(* IEC 61131-3 sources: stdmachine/plc/src/07_Tests, 6 files *)

(* ---- FB_AlarmManagerTest.st ---- *)
// Tests du gestionnaire d'alarmes (docs/04 § 10, docs/14 § 5)
FUNCTION_BLOCK FB_AlarmManagerTest EXTENDS TcUnit.FB_TestSuite
VAR
    stBuf : ST_AlarmBuffer;
END_VAR

RaiseTwiceOnce();
ClearedUnackedClosesOnAck();
LatchedEventClosesOnAck();
InfoClosesAtOnce();
AckedConditionClosesOnClear();

METHOD PRIVATE RaiseTwiceOnce
VAR
    fb : FB_AlarmManager;
END_VAR
TEST('RaiseTwiceOnce');
MEMSET(ADR(stBuf), 0, SIZEOF(stBuf));
fb.Bind(stBuf);
fb.Raise(1001, 101, 5, E_Severity.StationFault);
fb.Raise(1001, 101, 6, E_Severity.StationFault);
AssertEquals_UINT(Expected := 1, Actual := stBuf.nActive, Message := 'Une seule alarme pour la meme cle');
AssertEquals_UINT(Expected := 1, Actual := stBuf.aActive[1].nRepeat, Message := 'Repetition comptee');
AssertEquals_UDINT(Expected := 6, Actual := stBuf.aActive[1].nSubCode, Message := 'Sous-code mis a jour');
TEST_FINISHED();
END_METHOD

METHOD PRIVATE ClearedUnackedClosesOnAck
VAR
    fb : FB_AlarmManager;
END_VAR
TEST('ClearedUnackedClosesOnAck');
MEMSET(ADR(stBuf), 0, SIZEOF(stBuf));
fb.Bind(stBuf);
fb.Raise(2003, 100, 0, E_Severity.Warning);
fb.Clear(2003, 100);
AssertTrue(Condition := stBuf.nActive = 1 AND_THEN stBuf.aActive[1].eState = E_AlarmState.ClearedUnacked, Message := 'Disparue non acquittee : reste affichee');
fb.AckWarning(2003, 100, 'test');
AssertEquals_UINT(Expected := 0, Actual := stBuf.nActive, Message := 'Acquittee : close');
TEST_FINISHED();
END_METHOD

METHOD PRIVATE LatchedEventClosesOnAck
VAR
    fb : FB_AlarmManager;
END_VAR
TEST('LatchedEventClosesOnAck');
MEMSET(ADR(stBuf), 0, SIZEOF(stBuf));
fb.Bind(stBuf);
fb.RaiseEvent(1000, 901, 1, E_Severity.StationFault);
fb.AckFaults(1, FALSE, 'test');
AssertEquals_UINT(Expected := 0, Actual := stBuf.nActive, Message := 'Alarme sur evenement close a l acquittement');
TEST_FINISHED();
END_METHOD

METHOD PRIVATE InfoClosesAtOnce
VAR
    fb : FB_AlarmManager;
END_VAR
TEST('InfoClosesAtOnce');
MEMSET(ADR(stBuf), 0, SIZEOF(stBuf));
fb.Bind(stBuf);
fb.RaiseEvent(0, 916, 2, E_Severity.Info);
AssertEquals_UINT(Expected := 0, Actual := stBuf.nActive, Message := 'Information close des son apparition');
AssertEquals_UDINT(Expected := 2, Actual := stBuf.nWriteSeq, Message := 'Evenements apparition et cloture ecrits');
TEST_FINISHED();
END_METHOD

METHOD PRIVATE AckedConditionClosesOnClear
VAR
    fb : FB_AlarmManager;
END_VAR
TEST('AckedConditionClosesOnClear');
MEMSET(ADR(stBuf), 0, SIZEOF(stBuf));
fb.Bind(stBuf);
fb.Raise(3001, 100, 0, E_Severity.Warning);
fb.AckWarning(0, 0, 'test');
AssertTrue(Condition := stBuf.nActive = 1 AND_THEN stBuf.aActive[1].eState = E_AlarmState.ActiveAcked, Message := 'Acquittee, cause presente : reste active');
fb.Clear(3001, 100);
AssertEquals_UINT(Expected := 0, Actual := stBuf.nActive, Message := 'Cause disparue apres acquittement : close');
TEST_FINISHED();
END_METHOD
END_FUNCTION_BLOCK

(* ---- FB_HelpersTest.st ---- *)
// Tests des fonctions de base : CRC-32, comparaisons, opérations de SetVar, verdicts, états de calibration
FUNCTION_BLOCK FB_HelpersTest EXTENDS TcUnit.FB_TestSuite
VAR
END_VAR

Crc32Reference();
Crc32Incremental();
CompareTerms();
ApplyOperations();
VerdictOfData();
CalibStateRoundTrip();

METHOD PRIVATE Crc32Reference
VAR
    fb : FB_Crc32;
    s : STRING(20) := '123456789';
END_VAR
TEST('Crc32Reference');
fb.Begin(ADR(s), 9);
AssertTrue(Condition := fb.Step(1000), Message := 'Calcul termine en un pas');
AssertEquals_UDINT(Expected := 16#CBF43926, Actual := fb.Value, Message := 'CRC-32 IEEE de 123456789');
TEST_FINISHED();
END_METHOD

METHOD PRIVATE Crc32Incremental
VAR
    fb : FB_Crc32;
    s : STRING(20) := '123456789';
    n : INT;
END_VAR
TEST('Crc32Incremental');
fb.Begin(ADR(s), 9);
WHILE NOT fb.Step(2) AND n < 10 DO n := n + 1; END_WHILE
AssertEquals_INT(Expected := 4, Actual := n, Message := 'Cinq tranches de deux octets au plus');
AssertEquals_UDINT(Expected := 16#CBF43926, Actual := fb.Value, Message := 'Meme CRC par tranches');
TEST_FINISHED();
END_METHOD

METHOD PRIVATE CompareTerms
TEST('CompareTerms');
AssertTrue(Condition := F_Compare(1.0, E_Cmp.Eq, 1.0), Message := 'Eq');
AssertTrue(Condition := F_Compare(1.0, E_Cmp.Ne, 2.0), Message := 'Ne');
AssertTrue(Condition := F_Compare(1.0, E_Cmp.Lt, 2.0), Message := 'Lt');
AssertTrue(Condition := F_Compare(2.0, E_Cmp.Le, 2.0), Message := 'Le egal');
AssertFalse(Condition := F_Compare(2.0, E_Cmp.Gt, 2.0), Message := 'Gt strict');
AssertTrue(Condition := F_Compare(2.0, E_Cmp.Ge, 2.0), Message := 'Ge egal');
AssertTrue(Condition := F_Compare(1.0, E_Cmp.IsTrue, 0.0), Message := 'IsTrue');
AssertTrue(Condition := F_Compare(0.0, E_Cmp.IsFalse, 0.0), Message := 'IsFalse');
TEST_FINISHED();
END_METHOD

METHOD PRIVATE ApplyOperations
TEST('ApplyOperations');
AssertEquals_LREAL(Expected := 2.0, Actual := F_ApplyOp(5.0, 2.0, 0), Delta := 1.0E-9, Message := 'Affecter');
AssertEquals_LREAL(Expected := 7.0, Actual := F_ApplyOp(5.0, 2.0, 1), Delta := 1.0E-9, Message := 'Ajouter');
AssertEquals_LREAL(Expected := 3.0, Actual := F_ApplyOp(5.0, 2.0, 2), Delta := 1.0E-9, Message := 'Soustraire');
TEST_FINISHED();
END_METHOD

METHOD PRIVATE VerdictOfData
TEST('VerdictOfData');
AssertTrue(Condition := F_Verdict(0.0) = E_Verdict.Undefined, Message := '0 : non defini');
AssertTrue(Condition := F_Verdict(1.0) = E_Verdict.Good, Message := '1 : bon');
AssertTrue(Condition := F_Verdict(2.0) = E_Verdict.Bad, Message := '2 : mauvais');
TEST_FINISHED();
END_METHOD

METHOD PRIVATE CalibStateRoundTrip
TEST('CalibStateRoundTrip');
AssertTrue(Condition := F_CalibStateOf(F_CalibStateNum(E_CalibState.Valid)) = E_CalibState.Valid, Message := 'Valid');
AssertTrue(Condition := F_CalibStateOf(F_CalibStateNum(E_CalibState.Expired)) = E_CalibState.Expired, Message := 'Expired');
AssertTrue(Condition := F_CalibStateOf(F_CalibStateNum(E_CalibState.Failed)) = E_CalibState.Failed, Message := 'Failed');
AssertTrue(Condition := F_CalibStateOf(F_CalibStateNum(E_CalibState.Running)) = E_CalibState.Never, Message := 'Running restaure en Never');
TEST_FINISHED();
END_METHOD
END_FUNCTION_BLOCK

(* ---- FB_ObjectsSimTest.st ---- *)
// Tests d'objets en simulation (docs/04 § 14) : cas nominal, Abort pendant l'action, override 0 % puis reprise,
// paramètre invalide, action inconnue. Tests sur plusieurs cycles : l'état est gardé dans le bloc de test.
FUNCTION_BLOCK FB_ObjectsSimTest EXTENDS TcUnit.FB_TestSuite
VAR
    // Temporisation
    stCfgTimer : ST_ObjConfig;
    fbTimer : FB_Timer;
    stParTimer : ST_ActParams;
    nTimerStep : INT;
    fTimerMs : LREAL;
    // Vérin sans capteur
    stCfgCyl : ST_ObjConfig;
    fbCyl : FB_Cylinder;
    stParCyl : ST_ActParams;
    nCylStep : INT;
    fCylMs : LREAL;
    // Vérin interrompu
    stCfgCylAbort : ST_ObjConfig;
    fbCylAbort : FB_Cylinder;
    nAbortStep : INT;
    // Éclairage
    stCfgLight : ST_ObjConfig;
    fbLight : FB_Light;
    stParLight : ST_ActParams;
    nLightStep : INT;
    fLightMs : LREAL;
    // Magasin
    stCfgMag : ST_ObjConfig;
    fbMag : FB_Magazine;
    stParMag : ST_ActParams;
    nMagStep : INT;
END_VAR

TimerWaitsItsDuration();
CylinderOverrideZeroWaits();
CylinderAbortDuringMove();
LightFlashEnds();
MagazineCells();

METHOD PRIVATE _Cfg
VAR_IN_OUT
    stCfg : ST_ObjConfig;
END_VAR
VAR_INPUT
    nType : UINT;
    nLocalId : UINT;
END_VAR
MEMSET(ADR(stCfg), 0, SIZEOF(stCfg));
stCfg.nType := nType;
stCfg.nLocalId := nLocalId;
stCfg.nStableId := 1000 + nLocalId;
stCfg.sName := 'Essai';
stCfg.bSimulated := TRUE;
stCfg.fOverride := 100;
END_METHOD

METHOD PRIVATE TimerWaitsItsDuration
TEST('TimerWaitsItsDuration');
CASE nTimerStep OF
    0:
        _Cfg(stCfgTimer, GVL_Catalog.Type_Timer, 1);
        AssertTrue(Condition := fbTimer.Configure(refCfg := stCfgTimer, nStation := 1, nPoolIndex := 1, ipParent := 0, ipLocks := 0, ipAlarms := 0),
                   Message := 'Configuration acceptee');
        stParTimer.aKind[1] := E_ParamKind.Real;
        stParTimer.aReal[1] := 100;
        AssertTrue(Condition := fbTimer.Start(GVL_Catalog.Timer_Attendre, stParTimer, FALSE) = E_StartResult.Accepted, Message := 'Attendre accepte');
        nTimerStep := 1;
    1:
        fbTimer.Cycle();
        fTimerMs := fTimerMs + F_CycleMs();
        IF fbTimer.ActStatus = E_ActStatus.Done THEN
            AssertTrue(Condition := fTimerMs >= 95.0 AND fTimerMs <= 300.0, Message := 'Duree respectee');
            TEST_FINISHED();
            nTimerStep := 2;
        ELSIF fTimerMs > 2000.0 THEN
            AssertTrue(Condition := FALSE, Message := 'Attendre ne finit pas');
            TEST_FINISHED();
            nTimerStep := 2;
        END_IF
END_CASE
END_METHOD

// Override 0 % : le vérin ne part pas ; à 100 % il finit (docs/04 § 7.4)
METHOD PRIVATE CylinderOverrideZeroWaits
TEST('CylinderOverrideZeroWaits');
CASE nCylStep OF
    0:
        _Cfg(stCfgCyl, GVL_Catalog.Type_Cylinder, 2);
        stCfgCyl.aSignal[1].eKind := E_SignalKind.DO;
        stCfgCyl.aSignal[1].nIndex := 0;
        stCfgCyl.aParam[3] := 200;           // temps de mouvement sans capteur
        stCfgCyl.fOverride := 0;
        AssertTrue(Condition := fbCyl.Configure(refCfg := stCfgCyl, nStation := 1, nPoolIndex := 1, ipParent := 0, ipLocks := 0, ipAlarms := 0),
                   Message := 'Configuration acceptee');
        AssertTrue(Condition := fbCyl.Start(GVL_Catalog.Cylinder_MoveTravail, stParCyl, FALSE) = E_StartResult.Accepted, Message := 'Move travail accepte');
        nCylStep := 1;
    1:
        fbCyl.Cycle();
        fCylMs := fCylMs + F_CycleMs();
        IF fCylMs >= 500.0 THEN
            AssertTrue(Condition := fbCyl.ActStatus = E_ActStatus.Busy, Message := 'A 0 % le vérin attend');
            stCfgCyl.fOverride := 100;
            fCylMs := 0;
            nCylStep := 2;
        END_IF
    2:
        fbCyl.Cycle();
        fCylMs := fCylMs + F_CycleMs();
        IF fbCyl.ActStatus = E_ActStatus.Done OR fCylMs > 3000.0 THEN
            AssertTrue(Condition := fbCyl.ActStatus = E_ActStatus.Done, Message := 'Reprise a 100 % : fin du mouvement');
            TEST_FINISHED();
            nCylStep := 3;
        END_IF
END_CASE
END_METHOD

METHOD PRIVATE CylinderAbortDuringMove
TEST('CylinderAbortDuringMove');
CASE nAbortStep OF
    0:
        _Cfg(stCfgCylAbort, GVL_Catalog.Type_Cylinder, 3);
        stCfgCylAbort.aSignal[1].eKind := E_SignalKind.DO;
        stCfgCylAbort.aSignal[1].nIndex := 1;
        stCfgCylAbort.aParam[3] := 1000;
        fbCylAbort.Configure(refCfg := stCfgCylAbort, nStation := 1, nPoolIndex := 2, ipParent := 0, ipLocks := 0, ipAlarms := 0);
        fbCylAbort.Start(GVL_Catalog.Cylinder_MoveTravail, stParCyl, FALSE);
        nAbortStep := 1;
    1:
        fbCylAbort.Cycle();
        fbCylAbort.Abort();
        fbCylAbort.Cycle();                 // le statut est publié au cycle
        AssertTrue(Condition := fbCylAbort.ActStatus = E_ActStatus.Error, Message := 'Action interrompue');
        AssertEquals_UINT(Expected := GVL_Catalog.Err_Aborted, Actual := fbCylAbort.Status.nErrorCode, Message := 'Code Interrompue par Abort');
        AssertTrue(Condition := fbCylAbort.NodeState <> E_ObjState.Error, Message := 'Abort ne met pas l objet en erreur');
        AssertTrue(Condition := fbCylAbort.Start(9999, stParCyl, FALSE) = E_StartResult.UnknownAction, Message := 'Action inconnue refusee');
        TEST_FINISHED();
        nAbortStep := 2;
END_CASE
END_METHOD

METHOD PRIVATE LightFlashEnds
TEST('LightFlashEnds');
CASE nLightStep OF
    0:
        _Cfg(stCfgLight, GVL_Catalog.Type_Light, 4);
        stCfgLight.aSignal[1].eKind := E_SignalKind.DO;
        stCfgLight.aSignal[1].nIndex := 2;
        stCfgLight.aParam[2] := 80;
        stCfgLight.aParam[3] := 50;
        fbLight.Configure(refCfg := stCfgLight, nStation := 1, nPoolIndex := 1, ipParent := 0, ipLocks := 0, ipAlarms := 0);
        AssertTrue(Condition := fbLight.Start(GVL_Catalog.Light_Allumer, stParLight, FALSE) = E_StartResult.Accepted, Message := 'Allumer accepte');
        AssertTrue(Condition := fbLight.ActStatus = E_ActStatus.Done, Message := 'Allumer est immediat');
        AssertTrue(Condition := fbLight.Start(GVL_Catalog.Light_Flasher, stParLight, FALSE) = E_StartResult.Accepted, Message := 'Flasher accepte');
        nLightStep := 1;
    1:
        fbLight.Cycle();
        fLightMs := fLightMs + F_CycleMs();
        IF fbLight.ActStatus = E_ActStatus.Done OR fLightMs > 1000.0 THEN
            AssertTrue(Condition := fbLight.ActStatus = E_ActStatus.Done AND fLightMs >= 45.0, Message := 'Flash de 50 ms termine');
            AssertEquals_LREAL(Expected := 0.0, Actual := fbLight.Status.aValue[1], Delta := 0.0, Message := 'Eteint apres le flash');
            TEST_FINISHED();
            nLightStep := 2;
        END_IF
END_CASE
END_METHOD

METHOD PRIVATE MagazineCells
TEST('MagazineCells');
CASE nMagStep OF
    0:
        _Cfg(stCfgMag, GVL_Catalog.Type_Magazine, 5);
        stCfgMag.aSignal[1].eKind := E_SignalKind.DI;
        stCfgMag.aSignal[4].eKind := E_SignalKind.DO;
        stCfgMag.aSignal[4].nIndex := 3;
        stCfgMag.aSignal[5].eKind := E_SignalKind.DO;
        stCfgMag.aSignal[5].nIndex := 4;
        stCfgMag.aParam[1] := 2;            // 2 lignes
        stCfgMag.aParam[2] := 3;            // 3 colonnes
        stCfgMag.aParam[3] := 10;
        stCfgMag.aParam[4] := 20;
        fbMag.Configure(refCfg := stCfgMag, nStation := 1, nPoolIndex := 1, ipParent := 0, ipLocks := 0, ipAlarms := 0);
        fbMag.Start(GVL_Catalog.Magazine_PresenterPlateauSuivant, stParMag, FALSE);
        nMagStep := 1;
    1:
        fbMag.Cycle();
        IF fbMag.ActStatus <> E_ActStatus.Busy THEN
            AssertTrue(Condition := fbMag.ActStatus = E_ActStatus.Done, Message := 'Plateau presente en simulation');
            // Case 5 : ligne 2, colonne 2
            stParMag.aKind[1] := E_ParamKind.Real;
            stParMag.aReal[1] := 5;
            fbMag.Start(GVL_Catalog.Magazine_PositionDeLaCase, stParMag, FALSE);
            AssertEquals_LREAL(Expected := 10.0, Actual := fbMag.Results.stPos.fX, Delta := 1.0E-6, Message := 'X de la case 5');
            AssertEquals_LREAL(Expected := 20.0, Actual := fbMag.Results.stPos.fY, Delta := 1.0E-6, Message := 'Y de la case 5');
            stParMag.aReal[1] := 1;
            stParMag.aKind[2] := E_ParamKind.Real;
            stParMag.aReal[2] := 1;
            fbMag.Start(GVL_Catalog.Magazine_MarquerCase, stParMag, FALSE);
            stParMag.aReal[1] := 0;
            fbMag.Start(GVL_Catalog.Magazine_PositionDeLaCase, stParMag, FALSE);
            AssertEquals_LREAL(Expected := 2.0, Actual := fbMag.Results.aReal[2], Delta := 0.0, Message := 'Prochaine case libre : 2');
            fbMag.Start(GVL_Catalog.Magazine_LireOccupation, stParMag, FALSE);
            AssertEquals_LREAL(Expected := 1.0, Actual := fbMag.Results.aReal[1], Delta := 0.0, Message := 'Une case occupee');
            AssertEquals_LREAL(Expected := 5.0, Actual := fbMag.Results.aReal[2], Delta := 0.0, Message := 'Cinq cases libres');
            TEST_FINISHED();
            nMagStep := 2;
        END_IF
END_CASE
END_METHOD
END_FUNCTION_BLOCK

(* ---- FB_PackMLTest.st ---- *)
// Tests de la machine d'états PackML réduite (docs/05 § 2)
FUNCTION_BLOCK FB_PackMLTest EXTENDS TcUnit.FB_TestSuite
VAR
END_VAR

ResetThenIdle();
StartHoldRestart();
StopCompletes();
FaultAborts();
ClearReturnsStopped();
RejectedCommands();

METHOD PRIVATE ResetThenIdle
VAR
    fb : FB_PackML;
END_VAR
TEST('ResetThenIdle');
fb(eCmd := E_Cmd.Reset, bStateComplete := FALSE, bFault := FALSE);
AssertTrue(Condition := fb.eState = E_State.Resetting AND fb.bEntry, Message := 'Reset depuis Stopped : Resetting');
fb(eCmd := E_Cmd.None, bStateComplete := FALSE, bFault := FALSE);
AssertTrue(Condition := fb.eState = E_State.Resetting AND NOT fb.bEntry, Message := 'Resetting tant que le travail n est pas fini');
fb(eCmd := E_Cmd.None, bStateComplete := TRUE, bFault := FALSE);
AssertTrue(Condition := fb.eState = E_State.Idle, Message := 'Resetting termine : Idle');
TEST_FINISHED();
END_METHOD

METHOD PRIVATE StartHoldRestart
VAR
    fb : FB_PackML;
END_VAR
TEST('StartHoldRestart');
fb(eCmd := E_Cmd.Reset);
fb(eCmd := E_Cmd.None, bStateComplete := TRUE);
fb(eCmd := E_Cmd.Start, bStateComplete := FALSE);
AssertTrue(Condition := fb.eState = E_State.Execute, Message := 'Start depuis Idle : Execute');
fb(eCmd := E_Cmd.Hold);
AssertTrue(Condition := fb.eState = E_State.Held, Message := 'Hold : Held');
fb(eCmd := E_Cmd.Start);
AssertTrue(Condition := fb.eState = E_State.Execute, Message := 'Start depuis Held : Execute');
TEST_FINISHED();
END_METHOD

METHOD PRIVATE StopCompletes
VAR
    fb : FB_PackML;
END_VAR
TEST('StopCompletes');
fb(eCmd := E_Cmd.Reset);
fb(eCmd := E_Cmd.None, bStateComplete := TRUE);
fb(eCmd := E_Cmd.Start, bStateComplete := FALSE);
fb(eCmd := E_Cmd.Stop);
AssertTrue(Condition := fb.eState = E_State.Stopping, Message := 'Stop : Stopping');
fb(eCmd := E_Cmd.None, bStateComplete := TRUE);
AssertTrue(Condition := fb.eState = E_State.Stopped, Message := 'Stopping termine : Stopped');
TEST_FINISHED();
END_METHOD

METHOD PRIVATE FaultAborts
VAR
    fb : FB_PackML;
END_VAR
TEST('FaultAborts');
fb(eCmd := E_Cmd.Reset);
fb(eCmd := E_Cmd.None, bStateComplete := TRUE);
fb(eCmd := E_Cmd.Start, bStateComplete := FALSE);
fb(eCmd := E_Cmd.None, bFault := TRUE);
AssertTrue(Condition := fb.eState = E_State.Aborted, Message := 'Defaut en Execute : Aborted');
fb(eCmd := E_Cmd.Start, bFault := FALSE);
AssertTrue(Condition := fb.eState = E_State.Aborted, Message := 'Start refuse en Aborted');
TEST_FINISHED();
END_METHOD

METHOD PRIVATE ClearReturnsStopped
VAR
    fb : FB_PackML;
END_VAR
TEST('ClearReturnsStopped');
fb(eCmd := E_Cmd.Abort);
AssertTrue(Condition := fb.eState = E_State.Aborted, Message := 'Abort depuis Stopped : Aborted');
fb(eCmd := E_Cmd.Clear);
AssertTrue(Condition := fb.eState = E_State.Clearing, Message := 'Clear : Clearing');
fb(eCmd := E_Cmd.None, bStateComplete := TRUE);
AssertTrue(Condition := fb.eState = E_State.Stopped, Message := 'Clearing termine : Stopped');
TEST_FINISHED();
END_METHOD

METHOD PRIVATE RejectedCommands
VAR
    fb : FB_PackML;
END_VAR
TEST('RejectedCommands');
AssertFalse(Condition := fb.Accepts(E_Cmd.Start), Message := 'Start refuse en Stopped');
AssertFalse(Condition := fb.Accepts(E_Cmd.Hold), Message := 'Hold refuse en Stopped');
AssertTrue(Condition := fb.Accepts(E_Cmd.Reset), Message := 'Reset accepte en Stopped');
fb(eCmd := E_Cmd.Start);
AssertTrue(Condition := fb.eState = E_State.Stopped, Message := 'Start sans effet en Stopped');
TEST_FINISHED();
END_METHOD
END_FUNCTION_BLOCK

(* ---- FB_ScenarioEntryExitTest.st ---- *)
// Scénario de bout en bout (docs/05 § 12.1, docs/06 § 6.1) avec le système planaire simulé : une machine de deux
// stations (Chargement, rôle Entrée ; Déchargement, rôle Sortie), deux movers, un OF de 3 pièces.
// Déploiement par le handshake réel (zone d'attente, sommes de contrôle, Activate), OF, Reset, Start,
// puis arrêt automatique « OF terminé » avec 3 bonnes et aucune pièce sur les movers.
FUNCTION_BLOCK FB_ScenarioEntryExitTest EXTENDS TcUnit.FB_TestSuite
VAR
    fbMachine : FB_Machine;
    fbCrc : FB_Crc32;
    nStep : INT;
    fStepMs : LREAL;
    nSeq : UDINT;
    nOrder : UDINT;                 // n° d'OF propre à chaque exécution (les OF sont persistants)
    k : INT;
END_VAR

EntryExitThreeParts();

METHOD PRIVATE EntryExitThreeParts
VAR
    m : REFERENCE TO ST_MachineData;
    n : USINT;
END_VAR
TEST('EntryExitThreeParts');
IF nStep >= 100 THEN RETURN; END_IF
fbMachine();
fStepMs := fStepMs + F_CycleMs();
CASE nStep OF
    0:  // Zone d'attente
        MEMSET(ADR(GVL_Hmi.stStaging), 0, SIZEOF(GVL_Hmi.stStaging));
        m REF= GVL_Hmi.stStaging.stMachine;
        m.sMachineName := 'ESSAI';
        m.nMovers := 2;
        m.nSlots := 1;
        m.fOverride := 100;
        m.nNoStationMs := 60000;
        m.aGroup[1].bUsed := TRUE;
        m.aGroup[1].sName := 'Chargement';
        m.aGroup[1].eRole := E_GroupRole.Entry;
        m.aGroup[1].nStationMask := 1;
        m.aGroup[1].nOperations := 1;
        m.aGroup[1].nPriority := 5;
        m.aGroup[2].bUsed := TRUE;
        m.aGroup[2].sName := 'Dechargement';
        m.aGroup[2].eRole := E_GroupRole.Exit;
        m.aGroup[2].nStationMask := 2;
        m.aGroup[2].nOperations := 1;
        m.aGroup[2].nPriority := 5;
        FOR n := 1 TO 2 DO
            m.aStation[n].bUsed := TRUE;
            m.aStation[n].nGroupMask := SHL(UINT#1, n - 1);
            m.aStation[n].nWorkPos := n;
            m.aStation[n].fOverride := 100;
        END_FOR
        m.aStation[1].sName := 'Entree';
        m.aStation[2].sName := 'Sortie';
        m.nPlanarPos := 5;
        _PlanarPos(1, 100, 100, E_PlanarPosKind.Work, 1);
        _PlanarPos(2, 400, 100, E_PlanarPosKind.Work, 2);
        _PlanarPos(3, 100, 300, E_PlanarPosKind.Buffer, 0);
        _PlanarPos(4, 400, 300, E_PlanarPosKind.Buffer, 0);
        _PlanarPos(5, 700, 300, E_PlanarPosKind.Park, 0);
        m.nParkPos := 5;
        // Process général : Route(Chargement), Route(Déchargement), retour au début
        m.aTable[1].bUsed := TRUE;
        m.aTable[1].sName := 'Process general';
        m.aTable[1].eKind := E_TableKind.General;
        m.aTable[1].nStart := 1;
        m.aTable[1].nLength := 3;
        m.nInstrCount := 3;
        m.aInstr[1].eOp := E_Op.Route;
        m.aInstr[1].aArg[1] := 1;
        m.aInstr[1].aArg[2] := 1;
        m.aInstr[2].eOp := E_Op.Route;
        m.aInstr[2].aArg[1] := 2;
        m.aInstr[2].aArg[2] := 1;
        m.aInstr[3].eOp := E_Op.Jump;
        m.aInstr[3].aArg[1] := 1;
        // Chaque station : une opération (fonction n, opération 1) réduite à End(0)
        FOR n := 1 TO 2 DO
            GVL_Hmi.stStaging.aStation[n].aTable[1].bUsed := TRUE;
            GVL_Hmi.stStaging.aStation[n].aTable[1].sName := 'Operation';
            GVL_Hmi.stStaging.aStation[n].aTable[1].eKind := E_TableKind.Operation;
            GVL_Hmi.stStaging.aStation[n].aTable[1].nStart := 1;
            GVL_Hmi.stStaging.aStation[n].aTable[1].nLength := 1;
            GVL_Hmi.stStaging.aStation[n].nInstrCount := 1;
            GVL_Hmi.stStaging.aStation[n].aInstr[1].eOp := E_Op.End;
            GVL_Hmi.stStaging.aStation[n].nOpMapCount := 1;
            GVL_Hmi.stStaging.aStation[n].aOpMap[1].nGroup := n;
            GVL_Hmi.stStaging.aStation[n].aOpMap[1].nOperationNo := 1;
            GVL_Hmi.stStaging.aStation[n].aOpMap[1].nTable := 1;
        END_FOR
        // Sommes de contrôle, calculées comme la HMI le fera
        fbCrc.Begin(ADR(GVL_Hmi.stStaging.stMachine), SIZEOF(GVL_Hmi.stStaging.stMachine));
        fbCrc.Step(16#FFFFFFFF);
        GVL_Hmi.stDeploy.nCrcMachine := fbCrc.Value;
        FOR n := 1 TO GVL_Const.MAX_STATIONS DO
            fbCrc.Begin(ADR(GVL_Hmi.stStaging.aStation[n]), SIZEOF(GVL_Hmi.stStaging.aStation[n]));
            fbCrc.Step(16#FFFFFFFF);
            GVL_Hmi.stDeploy.aCrcStation[n] := fbCrc.Value;
        END_FOR
        fbCrc.Begin(ADR(GVL_Hmi.stStaging.aPressRecipe), SIZEOF(GVL_Hmi.stStaging.aPressRecipe));
        fbCrc.Step(16#FFFFFFFF);
        GVL_Hmi.stDeploy.nCrcRecipes := fbCrc.Value;
        GVL_Hmi.stDeploy.eCmd := E_DeployCmd.Activate;
        GVL_Hmi.stDeploy.nInstrSetRequired := 1;
        GVL_Hmi.stDeploy.nCatalogRequired := 1;
        GVL_Hmi.stDeploy.sUser := 'essai';
        nSeq := GVL_Hmi.stDeploy.nSeq + 1;
        GVL_Hmi.stDeploy.nSeq := nSeq;
        _Next(1);
    1:  // Réponse du déploiement
        IF GVL_Hmi.stDeployResp.nSeq = nSeq THEN
            AssertTrue(Condition := GVL_Hmi.stDeployResp.eResult = E_CmdResult.Accepted, Message := 'Deploiement accepte');
            AssertEquals_USINT(Expected := 0, Actual := GVL_Hmi.stDeployResp.nErrors, Message := 'Aucune erreur de deploiement');
            IF GVL_Hmi.stDeployResp.nErrors > 0 THEN
                AssertEquals_UINT(Expected := 0, Actual := GVL_Hmi.stDeployResp.aError[1].nCode, Message := 'Premiere erreur de deploiement');
            END_IF
            // OF de 3 pièces
            GVL_Hmi.stOrder.eCmd := E_OrderCmd.Activate;
            nOrder := LINT_TO_UDINT((F_NowUtc() / 10000000) MOD 1000000000) + 1;
            GVL_Hmi.stOrder.nOrder := nOrder;
            GVL_Hmi.stOrder.sNumber := 'OF-ESSAI';
            GVL_Hmi.stOrder.sReference := 'REF-1';
            GVL_Hmi.stOrder.nQuantity := 3;
            nSeq := GVL_Hmi.stOrder.nSeq + 1;
            GVL_Hmi.stOrder.nSeq := nSeq;
            _Next(2);
        ELSIF fStepMs > 5000 THEN
            _Abandon('Pas de reponse au deploiement');
        END_IF
    2:
        IF GVL_Hmi.stOrderResp.nSeq = nSeq THEN
            AssertTrue(Condition := GVL_Hmi.stOrderResp.eResult = E_CmdResult.Accepted, Message := 'OF accepte');
            _Command(E_Cmd.Reset);
            _Next(3);
        ELSIF fStepMs > 1000 THEN
            _Abandon('Pas de reponse a l OF');
        END_IF
    3:  // Reset : système planaire actif, movers détectés, stations Idle
        IF GVL_Hmi.stMachineStatus.eState = E_State.Idle THEN
            _Command(E_Cmd.Start);
            _Next(4);
        ELSIF fStepMs > 10000 THEN
            _Abandon('La machine n arrive pas en Idle');
        END_IF
    4:
        IF GVL_Hmi.stMachineStatus.eState = E_State.Execute THEN
            _Next(5);
        ELSIF fStepMs > 1000 THEN
            _Abandon('La machine ne demarre pas');
        END_IF
    5:  // Production jusqu'à l'arrêt automatique « OF terminé »
        IF GVL_Hmi.stMachineStatus.eState = E_State.Stopped THEN
            AssertTrue(Condition := GVL_Hmi.stMachineStatus.eStopReason = E_StopReason.OrderComplete, Message := 'Arret automatique OF termine');
            AssertEquals_UINT(Expected := 0, Actual := GVL_Hmi.stMachineStatus.nPartsInProcess, Message := 'Aucune piece sur les movers');
            FOR k := 1 TO GVL_Const.MAX_ORDERS DO
                IF GVL_Hmi.stMachineStatus.aOrder[k].nOrder = nOrder THEN
                    AssertEquals_UDINT(Expected := 3, Actual := GVL_Hmi.stMachineStatus.aOrder[k].nGood, Message := 'Trois bonnes');
                    AssertEquals_UDINT(Expected := 0, Actual := GVL_Hmi.stMachineStatus.aOrder[k].nBad, Message := 'Aucune mauvaise');
                    AssertTrue(Condition := GVL_Hmi.stMachineStatus.aOrder[k].eState = E_OrderState.Done, Message := 'OF termine');
                END_IF
            END_FOR
            AssertTrue(Condition := GVL_Hmi.stTraces.nWriteSeq >= 6, Message := 'Une trace par operation et par piece');
            TEST_FINISHED();
            nStep := 100;
        ELSIF GVL_Hmi.stMachineStatus.eState = E_State.Aborted THEN
            _Abandon('La machine est passee Aborted');
        ELSIF fStepMs > 60000 THEN
            _Abandon('L OF ne se termine pas en 60 s');
        END_IF
END_CASE
END_METHOD

METHOD PRIVATE _PlanarPos
VAR_INPUT
    nIndex : INT;
    fX : LREAL;
    fY : LREAL;
    eKind : E_PlanarPosKind;
    nStation : USINT;
END_VAR
GVL_Hmi.stStaging.stMachine.aPlanarPos[nIndex].stPos.fX := fX;
GVL_Hmi.stStaging.stMachine.aPlanarPos[nIndex].stPos.fY := fY;
GVL_Hmi.stStaging.stMachine.aPlanarPos[nIndex].eKind := eKind;
GVL_Hmi.stStaging.stMachine.aPlanarPos[nIndex].nStation := nStation;
END_METHOD

METHOD PRIVATE _Command
VAR_INPUT
    eCmd : E_Cmd;
END_VAR
GVL_Hmi.stCmd.nTarget := 0;
GVL_Hmi.stCmd.bSetMode := FALSE;
GVL_Hmi.stCmd.eCmd := eCmd;
GVL_Hmi.stCmd.sUser := 'essai';
GVL_Hmi.stCmd.nSeq := GVL_Hmi.stCmd.nSeq + 1;
END_METHOD

METHOD PRIVATE _Next
VAR_INPUT
    nNext : INT;
END_VAR
nStep := nNext;
fStepMs := 0;
END_METHOD

METHOD PRIVATE _Fail
VAR_INPUT
    sWhy : STRING(80);
END_VAR
AssertTrue(Condition := FALSE, Message := sWhy);
TEST_FINISHED();
nStep := 100;
END_METHOD
END_FUNCTION_BLOCK

(* ---- PRG_StdMachineTests.st ---- *)
// Programme de test TcUnit (docs/04 § 14) : à appeler dans la tâche du projet de test, qui référence
// StdMachineLib et TcUnit. Chaque suite déclarée ici est exécutée par TcUnit.RUN().
PROGRAM PRG_StdMachineTests
VAR
    fbPackML : FB_PackMLTest;
    fbHelpers : FB_HelpersTest;
    fbAlarms : FB_AlarmManagerTest;
    fbObjects : FB_ObjectsSimTest;
    fbScenario : FB_ScenarioEntryExitTest;
END_VAR

TcUnit.RUN();
END_PROGRAM
